(* IEC 61131-3 sources: Codesys_IAP/Demo/PLC1/Magazijn Overzetter Simulatie Structured Text 2V1_tekst/Programma Structured Text/States, 3 files *)

(* ---- magazijnStates.st ---- *)
(*#### DECLARATIE ####*)
// Datum : 17 december 2020, Auteur: Gerard Harkema
{attribute 'qualified_only'}
{attribute 'strict'}
TYPE magazijnStates :
(
	idle := 0,
	in,
	travel_out,
	out,
	travel_in,
	error
);
END_TYPE

(* ---- overzetterStates.st ---- *)
(*#### DECLARATIE ####*)
// Datum : 17 december 2020, Auteur: Gerard Harkema
{attribute 'qualified_only'}
{attribute 'strict'}
TYPE overzetterStates :
(
	idle := 0,
	is_links,
	vaccuum_aanzetten,
	ga_naar_rechts,
	is_rechts,
	vaccuum_lossen,
	ga_naar_midden,
	is_midden,
	ga_naar_links,
	error
);
END_TYPE

(* ---- stationStates.st ---- *)
(*#### DECLARATIE ####*)
// Datum : 26 november 2026, Auteur: Gerard Harkema
{attribute 'qualified_only'}
{attribute 'strict'}
TYPE stationStates :
(
	idle := 0,
	magazijn_uitstoten,
	wacht_magazijn_klaar,
	overzetten,
	wacht_overzetter_klaar,
	error
);
END_TYPE
